FUNCTION_BLOCK SortingSafeServices (* Existing ownership, command and measured home conditions. *)
  (* Standard: 61499-2 *)
  (* Version 3.0, 2026-11-12, sorting2n, sorting2n *)
  PACKAGE Main;
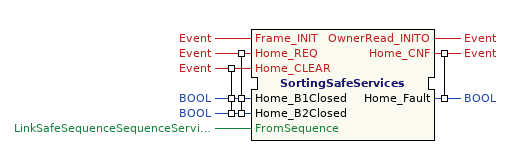
  EVENT_INPUT
    Frame_INIT;
    Home_REQ WITH Home_B1Closed, Home_B2Closed;
    Home_CLEAR WITH Home_B1Closed, Home_B2Closed;
  END_EVENT
  EVENT_OUTPUT
    OwnerRead_INITO;
    Home_CNF WITH Home_Fault;
  END_EVENT
  VAR_INPUT
    Home_B1Closed : BOOL;
    Home_B2Closed : BOOL;
  END_VAR
  VAR_OUTPUT
    Home_Fault : BOOL;
  END_VAR
  SOCKETS
    FromSequence : LinkSafeSequenceSequenceServices;
  END_SOCKETS
  FBS
    Frame : SortingCommandFrame;
    Ownership : SortingOwnership;
    OwnerRead : SYMLINKMULTIVARDST(QI := TRUE, NAME1 := '$${PATH:4}Conveyor.sc.progLocal', NAME2 := '$${PATH:4}Branch1.sc.progLocal', NAME3 := '$${PATH:4}Branch2.sc.progLocal', NAME4 := '$${PATH:4}Stopper.sc.progLocal'); {SET_ATTRIBUTE(Configuration.GenericFBType.InterfaceParams, Runtime.System#I:=4;VALUE${I$}:VTQBOOL,VTQBOOL,VTQBOOL,VTQBOOL)}
    OwnerWrite : SYMLINKMULTIVARSRC(QI := TRUE, NAME1 := '$${PATH:4}Conveyor.sc.progLocalSel', NAME2 := '$${PATH:4}Branch1.sc.progLocalSel', NAME3 := '$${PATH:4}Branch2.sc.progLocalSel', NAME4 := '$${PATH:4}Stopper.sc.progLocalSel'); {SET_ATTRIBUTE(Configuration.GenericFBType.InterfaceParams, Runtime.System#I:=4;VALUE${I$}:VTQBOOL,VTQBOOL,VTQBOOL,VTQBOOL)}
    WriteCommands : SYMLINKMULTIVARSRC(QI := TRUE, NAME1 := '$${PATH:4}Conveyor.sc.lsp', NAME2 := '$${PATH:4}Branch1.sc.lsp', NAME3 := '$${PATH:4}Branch2.sc.lsp', NAME4 := '$${PATH:4}Stopper.sc.lsp'); {SET_ATTRIBUTE(Configuration.GenericFBType.InterfaceParams, Runtime.System#I:=4;VALUE${I$}:VTQINT,VTQINT,VTQINT,VTQINT)}
    Home : SortingHomeConditions;
  END_FBS
  EVENT_CONNECTIONS
    Frame_INIT TO Frame.3E51AF3DA95F41C9;
    Frame.91A08A19905E4AC8 TO WriteCommands.INIT;
    WriteCommands.INITO TO Ownership.D514169649844923;
    Ownership.4CD8C065E39641C9 TO OwnerWrite.INIT;
    OwnerWrite.INITO TO OwnerRead.INIT;
    Ownership.B3E6986DDAA841AB TO OwnerWrite.REQ;
    OwnerRead.CNF TO Ownership.6D56496F53D1499B;
    OwnerRead.INITO TO Ownership.6D56496F53D1499B;
    Frame.FEDD90899323480E TO WriteCommands.REQ;
    Home_REQ TO Home.F4871D28B0594017;
    OwnerRead.INITO TO Home.CE64267AAD124F8D;
    Home.C188F07096974982 TO FromSequence.199423B8E3EA424D;
    OwnerRead.INITO TO OwnerRead_INITO;
    Home.199DF02180EA4007 TO Home_CNF;
    Home_CLEAR TO Home.27094514BA434C7A;
    FromSequence.011CF67C6620420F TO Ownership.8B11DD0F57C44878;
    Ownership.556ECCED2B7E4FE4 TO FromSequence.8705939D5B1442EC;
    FromSequence.A7B722B3D101427D TO Frame.B00E6A8BE1EB4052;
    FromSequence.8F745BA862BE446D TO Home.C8FE616D2B744827;
    FromSequence.DE074F0018CA41B7 TO Home.858AFA5821D243F1;
    Home.199DF02180EA4007 TO FromSequence.F3737632F0674E5B;
  END_CONNECTIONS
  DATA_CONNECTIONS
    OwnerRead.VALUE1 TO Ownership.3633AFB15F0E4D29;
    Ownership.AB3AFA1E5DB542BD TO OwnerWrite.VALUE1;
    OwnerRead.VALUE2 TO Ownership.AFBF64D6B6724875;
    Ownership.AB3AFA1E5DB542BD TO OwnerWrite.VALUE2;
    OwnerRead.VALUE3 TO Ownership.C6BAC61A3B114656;
    Ownership.AB3AFA1E5DB542BD TO OwnerWrite.VALUE3;
    OwnerRead.VALUE4 TO Ownership.0CBD0A2278FC4256;
    Ownership.AB3AFA1E5DB542BD TO OwnerWrite.VALUE4;
    Frame.1BE4F90CA0DE4A12 TO WriteCommands.VALUE1;
    Frame.E7BCFB58D0E944F4 TO WriteCommands.VALUE2;
    Frame.FD5B17DC6BEA4636 TO WriteCommands.VALUE3;
    Frame.9F87DE883B874F73 TO WriteCommands.VALUE4;
    Home_B1Closed TO Home.6DF2726E50AE4D83;
    Home_B2Closed TO Home.305FF7EA37BC4E0C;
    Home.74C9C2C856054ACB TO Home_Fault;
    Ownership.3DD7BBA990934FB9 TO FromSequence.B0172C60E5884E40;
    Home.097D9CE53785454A TO FromSequence.A973A7B0624E4A64;
  END_CONNECTIONS
END_FUNCTION_BLOCK
